(* PLC project Vn_jump_cond, Beckhoff Automation GmbH TwinCAT PLC Control 3.5.13.21 *)
(* stored: creationDateTime 1970-01-01T00:00:00 *)

PROGRAM Vn_jump_cond

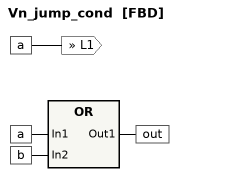
(* FBD diagram, written out as Structured Text *)
IF a THEN JMP L1; END_IF;
out := a OR b;
END_PROGRAM
